Fanuc KAREL source: ke00001.KL

-- PROVISIONAL review KL for V770-1; original PC SHA256 74a213ce18f14c7b02404300e3452b8ecbf02d11cbf0e1c1aedadeaa66ddea23
-- Incomplete behavior may be omitted. Consult companion uncertainty JSON. Do not deploy.
PROGRAM KE00001
%NOLOCKGROUP
BEGIN
  -- UNRESOLVED_PC offsets 5-12; opcodes 9D,23
  -- UNRESOLVED_PC offsets 17-41; opcodes 27,22,22,2A,22,31
  -- UNRESOLVED_PC offsets 46-50; opcodes 7F
END KE00001
